                                     Light_Guard_Bypass=>"Light_Guard_Bypass(1)",
                                     System_Busy:="System_1_Busy");
                100401:
                    "Feed_BCNV_Cnv1(1)"( System_No := 1,
                                     Level := 4,
                                     Light_Guard_IO:="LIGHT GUARDS C1101 - CH1",
                                     Light_Guard_Bypass=>"Light_Guard_Bypass(1)",
                                     System_Busy:="System_1_Busy");
                100501:
                    "Feed_BCNV_Cnv1(1)"( System_No := 1,
                                     Level := 5,
                                     Light_Guard_IO:="LIGHT GUARDS C1101 - CH1",
                                     Light_Guard_Bypass=>"Light_Guard_Bypass(1)",
                                     System_Busy:="System_1_Busy");
                100601:
                    "Feed_BCNV_Cnv1(1)"( System_No := 1,
                                     Level := 6,
                                     Light_Guard_IO:="LIGHT GUARDS C1101 - CH1",
                                     Light_Guard_Bypass=>"Light_Guard_Bypass(1)",
                                     System_Busy:="System_1_Busy");
                100701:
                    "Feed_BCNV_Cnv1(1)"( System_No := 1,
                                     Level := 7,
                                     Light_Guard_IO:="LIGHT GUARDS C1101 - CH1",
                                     Light_Guard_Bypass=>"Light_Guard_Bypass(1)",
                                     System_Busy:="System_1_Busy");
                100801:
                    "Feed_BCNV_Cnv1(1)"( System_No := 1,
                                     Level := 8,
                                     Light_Guard_IO:="LIGHT GUARDS C1101 - CH1",
                                     Light_Guard_Bypass=>"Light_Guard_Bypass(1)",
                                     System_Busy:="System_1_Busy");
                    //CNV 2
                110101:
                    "Feed_BCNV_Cnv2(1)"( System_No := 1,
                                     Level := 1,
                                     Light_Guard_IO:="LIGHT GUARDS C1201 - CH1",
                                     Light_Guard_Bypass=>"Light_Guard_Bypass(1)",
                                     System_Busy:="System_1_Busy");
                110201:
                    "Feed_BCNV_Cnv2(1)"( System_No := 1,
                                     Level := 2,
                                     Light_Guard_IO:="LIGHT GUARDS C1201 - CH1",
                                     Light_Guard_Bypass=>"Light_Guard_Bypass(1)",
                                     System_Busy:="System_1_Busy");
                110301:
                    "Feed_BCNV_Cnv2(1)"( System_No := 1,
                                     Level := 3,
                                     Light_Guard_IO:="LIGHT GUARDS C1201 - CH1",
                                     Light_Guard_Bypass=>"Light_Guard_Bypass(1)",
                                     System_Busy:="System_1_Busy");
                110401:
                    "Feed_BCNV_Cnv2(1)"( System_No := 1,
                                     Level := 4,
                                     Light_Guard_IO:="LIGHT GUARDS C1201 - CH1",
                                     Light_Guard_Bypass=>"Light_Guard_Bypass(1)",
                                     System_Busy:="System_1_Busy");
                110501:
                    "Feed_BCNV_Cnv2(1)"( System_No := 1,
                                     Level := 5,
                                     Light_Guard_IO:="LIGHT GUARDS C1201 - CH1",
                                     Light_Guard_Bypass=>"Light_Guard_Bypass(1)",
                                     System_Busy:="System_1_Busy");
                110601:
                    "Feed_BCNV_Cnv2(1)"( System_No := 1,
                                     Level := 6,
                                     Light_Guard_IO:="LIGHT GUARDS C1201 - CH1",
                                     Light_Guard_Bypass=>"Light_Guard_Bypass(1)",
                                     System_Busy:="System_1_Busy");
                110701:
                    "Feed_BCNV_Cnv2(1)"( System_No := 1,
                                     Level := 7,
                                     Light_Guard_IO:="LIGHT GUARDS C1201 - CH1",
                                     Light_Guard_Bypass=>"Light_Guard_Bypass(1)",
                                     System_Busy:="System_1_Busy");
                110801:
                    "Feed_BCNV_Cnv2(1)"( System_No := 1,
                                     Level := 8,
                                     Light_Guard_IO:="LIGHT GUARDS C1201 - CH1",
                                     Light_Guard_Bypass=>"Light_Guard_Bypass(1)",
                                     System_Busy:="System_1_Busy");
                    //SYSTEM 2
                    //CNV 1
                100102:
                    "Feed_BCNV_Cnv1(1)"(System_No := 2,
                                        Level := 1,
                                        Light_Guard_IO := "LIGHT GUARDS C2101 - CH1",
                                        Light_Guard_Bypass=>"Light_Guard_Bypass(2)",
                                        System_Busy := "System_2_Busy");
                100202:
                    "Feed_BCNV_Cnv1(1)"( System_No := 2,
                                     Level := 2,
                                     Light_Guard_IO:="LIGHT GUARDS C2101 - CH1",
                                     Light_Guard_Bypass=>"Light_Guard_Bypass(2)",
                                     System_Busy:="System_2_Busy");
                100302:
                    "Feed_BCNV_Cnv1(1)"( System_No := 2,
                                     Level := 3,
                                     Light_Guard_IO:="LIGHT GUARDS C2101 - CH1",
                                     Light_Guard_Bypass=>"Light_Guard_Bypass(2)",
                                     System_Busy:="System_2_Busy");
                100402:
                    "Feed_BCNV_Cnv1(1)"( System_No := 2,
                                     Level := 4,
                                     Light_Guard_IO:="LIGHT GUARDS C2101 - CH1",
                                     Light_Guard_Bypass=>"Light_Guard_Bypass(2)",
                                     System_Busy:="System_2_Busy");
                100502:
                    "Feed_BCNV_Cnv1(1)"( System_No := 2,
                                     Level := 5,
                                     Light_Guard_IO:="LIGHT GUARDS C2101 - CH1",
                                     Light_Guard_Bypass=>"Light_Guard_Bypass(2)",
                                     System_Busy:="System_2_Busy");
                100602:
                    "Feed_BCNV_Cnv1(1)"( System_No := 2,
                                     Level := 6,
                                     Light_Guard_IO:="LIGHT GUARDS C2101 - CH1",
                                     Light_Guard_Bypass=>"Light_Guard_Bypass(2)",
                                     System_Busy:="System_2_Busy");
                100702:
                    "Feed_BCNV_Cnv1(1)"( System_No := 2,
                                     Level := 7,
                                     Light_Guard_IO:="LIGHT GUARDS C2101 - CH1",
                                     Light_Guard_Bypass=>"Light_Guard_Bypass(2)",
                                     System_Busy:="System_2_Busy");
                100802:
                    "Feed_BCNV_Cnv1(1)"( System_No := 2,
                                     Level := 8,
                                     Light_Guard_IO:="LIGHT GUARDS C2101 - CH1",
                                     Light_Guard_Bypass=>"Light_Guard_Bypass(2)",
                                     System_Busy:="System_2_Busy");
                    //CNV 2
                110102:
                    "Feed_BCNV_Cnv2(1)"( System_No := 2,
                                     Level := 1,
                                     Light_Guard_IO:="LIGHT GUARDS C2201 - CH1",
                                     Light_Guard_Bypass=>"Light_Guard_Bypass(2)",
                                     System_Busy:="System_2_Busy");
                110202:
                    "Feed_BCNV_Cnv2(1)"( System_No := 2,
                                     Level := 2,
                                     Light_Guard_IO:="LIGHT GUARDS C2201 - CH1",
                                     Light_Guard_Bypass=>"Light_Guard_Bypass(2)",
                                     System_Busy:="System_2_Busy");
                110302:
                    "Feed_BCNV_Cnv2(1)"( System_No := 2,
                                     Level := 3,
                                     Light_Guard_IO:="LIGHT GUARDS C2201 - CH1",
                                     Light_Guard_Bypass=>"Light_Guard_Bypass(2)",
                                     System_Busy:="System_2_Busy");
                110402:
                    "Feed_BCNV_Cnv2(1)"( System_No := 2,
                                     Level := 4,
                                     Light_Guard_IO:="LIGHT GUARDS C2201 - CH1",
                                     Light_Guard_Bypass=>"Light_Guard_Bypass(2)",
                                     System_Busy:="System_2_Busy");
                110502:
                    "Feed_BCNV_Cnv2(1)"( System_No := 2,
                                     Level := 5,
                                     Light_Guard_IO:="LIGHT GUARDS C2201 - CH1",
                                     Light_Guard_Bypass=>"Light_Guard_Bypass(2)",
                                     System_Busy:="System_2_Busy");
                110602:
                    "Feed_BCNV_Cnv2(1)"( System_No := 2,
                                     Level := 6,
                                     Light_Guard_IO:="LIGHT GUARDS C2201 - CH1",
                                     Light_Guard_Bypass=>"Light_Guard_Bypass(2)",
                                     System_Busy:="System_2_Busy");
                110702:
                    "Feed_BCNV_Cnv2(1)"( System_No := 2,
                                     Level := 7,
                                     Light_Guard_IO:="LIGHT GUARDS C2201 - CH1",
                                     Light_Guard_Bypass=>"Light_Guard_Bypass(2)",
                                     System_Busy:="System_2_Busy");
                110802:
                    "Feed_BCNV_Cnv2(1)"( System_No := 2,
                                     Level := 8,
                                     Light_Guard_IO:="LIGHT GUARDS C2201 - CH1",
                                     Light_Guard_Bypass=>"Light_Guard_Bypass(2)",
                                     System_Busy:="System_2_Busy");
                    //SYSTEM 3
                    //CNV 1
                100103:
                    "Feed_BCNV_Cnv1(1)"( System_No := 3,
                                     Level := 1,
                                     Light_Guard_IO:="LIGHT GUARDS C3101 - CH1",
                                     Light_Guard_Bypass=>"Light_Guard_Bypass(3)",
                                     System_Busy:="System_3_Busy");
                100203:
                    "Feed_BCNV_Cnv1(1)"( System_No := 3,
                                     Level := 2,
                                     Light_Guard_IO:="LIGHT GUARDS C3101 - CH1",
                                     Light_Guard_Bypass=>"Light_Guard_Bypass(3)",
                                     System_Busy:="System_3_Busy");
                100303:
                    "Feed_BCNV_Cnv1(1)"( System_No := 3,
                                     Level := 3,
                                     Light_Guard_IO:="LIGHT GUARDS C3101 - CH1",
                                     Light_Guard_Bypass=>"Light_Guard_Bypass(3)",
                                     System_Busy:="System_3_Busy");
                100403:
                    "Feed_BCNV_Cnv1(1)"( System_No := 3,
                                     Level := 4,
                                     Light_Guard_IO:="LIGHT GUARDS C3101 - CH1",
                                     Light_Guard_Bypass=>"Light_Guard_Bypass(3)",
                                     System_Busy:="System_3_Busy");
                100503:
                    "Feed_BCNV_Cnv1(1)"( System_No := 3,
                                     Level := 5,
                                     Light_Guard_IO:="LIGHT GUARDS C3101 - CH1",
                                     Light_Guard_Bypass=>"Light_Guard_Bypass(3)",
                                     System_Busy:="System_3_Busy");
                100603:
                    "Feed_BCNV_Cnv1(1)"( System_No := 3,
                                     Level := 6,
                                     Light_Guard_IO:="LIGHT GUARDS C3101 - CH1",
                                     Light_Guard_Bypass=>"Light_Guard_Bypass(3)",
                                     System_Busy:="System_3_Busy");
                100703:
                    "Feed_BCNV_Cnv1(1)"( System_No := 3,
                                     Level := 7,
                                     Light_Guard_IO:="LIGHT GUARDS C3101 - CH1",
                                     Light_Guard_Bypass=>"Light_Guard_Bypass(3)",
                                     System_Busy:="System_3_Busy");
                100803:
                    "Feed_BCNV_Cnv1(1)"( System_No := 3,
                                     Level := 8,
                                     Light_Guard_IO:="LIGHT GUARDS C3101 - CH1",
                                     Light_Guard_Bypass=>"Light_Guard_Bypass(3)",
                                     System_Busy:="System_3_Busy");
                    //CNV 2
                110103:
                    "Feed_BCNV_Cnv2(1)"( System_No := 3,
                                     Level := 1,
                                     Light_Guard_IO:="LIGHT GUARDS C3201 - CH1",
                                     Light_Guard_Bypass=>"Light_Guard_Bypass(3)",
                                     System_Busy:="System_3_Busy");
                110203:
                    "Feed_BCNV_Cnv2(1)"( System_No := 3,
                                     Level := 2,
                                     Light_Guard_IO:="LIGHT GUARDS C3201 - CH1",
                                     Light_Guard_Bypass=>"Light_Guard_Bypass(3)",
                                     System_Busy:="System_3_Busy");
                110303:
                    "Feed_BCNV_Cnv2(1)"( System_No := 3,
                                     Level := 3,
                                     Light_Guard_IO:="LIGHT GUARDS C3201 - CH1",
                                     Light_Guard_Bypass=>"Light_Guard_Bypass(3)",
                                     System_Busy:="System_3_Busy");
                110403:
                    "Feed_BCNV_Cnv2(1)"( System_No := 3,
                                     Level := 4,
                                     Light_Guard_IO:="LIGHT GUARDS C3201 - CH1",
                                     Light_Guard_Bypass=>"Light_Guard_Bypass(3)",
                                     System_Busy:="System_3_Busy");
                110503:
                    "Feed_BCNV_Cnv2(1)"( System_No := 3,
                                     Level := 5,
                                     Light_Guard_IO:="LIGHT GUARDS C3201 - CH1",
                                     Light_Guard_Bypass=>"Light_Guard_Bypass(3)",
                                     System_Busy:="System_3_Busy");
                110603:
                    "Feed_BCNV_Cnv2(1)"( System_No := 3,
                                     Level := 6,
                                     Light_Guard_IO:="LIGHT GUARDS C3201 - CH1",
                                     Light_Guard_Bypass=>"Light_Guard_Bypass(3)",
                                     System_Busy:="System_3_Busy");
                110703:
                    "Feed_BCNV_Cnv2(1)"( System_No := 3,
                                     Level := 7,
                                     Light_Guard_IO:="LIGHT GUARDS C3201 - CH1",
                                     Light_Guard_Bypass=>"Light_Guard_Bypass(3)",
                                     System_Busy:="System_3_Busy");
                110803:
                    "Feed_BCNV_Cnv2(1)"( System_No := 3,
                                     Level := 8,
                                     Light_Guard_IO:="LIGHT GUARDS C3201 - CH1",
                                     Light_Guard_Bypass=>"Light_Guard_Bypass(3)",
                                     System_Busy:="System_3_Busy");
                    //SYSTEM 4
                    //CNV 2
                100104:
                    "Feed_BCNV_Cnv1(1)"( System_No := 4,
                                     Level := 1,
                                     Light_Guard_IO:=TRUE,
                                     Light_Guard_Bypass=>#No_Light_Guard,
                                     System_Busy:="System_4_Busy");
                100204:
                    "Feed_BCNV_Cnv1(1)"( System_No := 4,
                                     Level := 2,
                                     Light_Guard_IO:=TRUE,
                                     Light_Guard_Bypass=>#No_Light_Guard,
                                     System_Busy:="System_4_Busy");
                100304:
                    "Feed_BCNV_Cnv1(1)"( System_No := 4,
                                     Level := 3,
                                     Light_Guard_IO:=TRUE,
                                     Light_Guard_Bypass=>#No_Light_Guard,
                                     System_Busy:="System_4_Busy");
                100404:
                    "Feed_BCNV_Cnv1(1)"( System_No := 4,
                                     Level := 4,
                                     Light_Guard_IO:=TRUE,
                                     Light_Guard_Bypass=>#No_Light_Guard,
                                     System_Busy:="System_4_Busy");
                100504:
                    "Feed_BCNV_Cnv1(1)"( System_No := 4,
                                     Level := 5,
                                     Light_Guard_IO:=TRUE,
                                     Light_Guard_Bypass=>#No_Light_Guard,
                                     System_Busy:="System_4_Busy");
                100604:
                    "Feed_BCNV_Cnv1(1)"( System_No := 4,
                                     Level := 6,
                                     Light_Guard_IO:=TRUE,
                                     Light_Guard_Bypass=>#No_Light_Guard,
                                     System_Busy:="System_4_Busy");
                100704:
                    "Feed_BCNV_Cnv1(1)"( System_No := 4,
                                     Level := 7,
                                     Light_Guard_IO:=TRUE,
                                     Light_Guard_Bypass=>#No_Light_Guard,
                                     System_Busy:="System_4_Busy");
                100804:
                    "Feed_BCNV_Cnv1(1)"( System_No := 4,
                                     Level := 8,
                                     Light_Guard_IO:=TRUE,
                                     Light_Guard_Bypass=>#No_Light_Guard,
                                     System_Busy:="System_4_Busy");
                    //SYSTEM 5
                120005:
                    "Feed_ECNV(1)"( System_No := 5);
                    //CNV 2
                100105:
                    "Feed_BCNV_Cnv1(1)"( System_No := 5,
                                     Level := 1,
                                     Light_Guard_IO:=TRUE,
                                     Light_Guard_Bypass=>#No_Light_Guard,
                                     System_Busy:="System_5_Busy");
                100205:
                    "Feed_BCNV_Cnv1(1)"( System_No := 5,
                                     Level := 2,
                                     Light_Guard_IO:=TRUE,
                                     Light_Guard_Bypass=>#No_Light_Guard,
                                     System_Busy:="System_5_Busy");
                100305:
                    "Feed_BCNV_Cnv1(1)"( System_No := 5,
                                     Level := 3,
                                     Light_Guard_IO:=TRUE,
                                     Light_Guard_Bypass=>#No_Light_Guard,
                                     System_Busy:="System_5_Busy");
                100405:
                    "Feed_BCNV_Cnv1(1)"( System_No := 5,
                                     Level := 4,
                                     Light_Guard_IO:=TRUE,
                                     Light_Guard_Bypass=>#No_Light_Guard,
                                     System_Busy:="System_5_Busy");
                100505:
                    "Feed_BCNV_Cnv1(1)"( System_No := 5,
                                     Level := 5,
                                     Light_Guard_IO:=TRUE,
                                     Light_Guard_Bypass=>#No_Light_Guard,
                                     System_Busy:="System_5_Busy");
                100605:
                    "Feed_BCNV_Cnv1(1)"( System_No := 5,
                                     Level := 6,
                                     Light_Guard_IO:=TRUE,
                                     Light_Guard_Bypass=>#No_Light_Guard,
                                     System_Busy:="System_5_Busy");
                100705:
                    "Feed_BCNV_Cnv1(1)"( System_No := 5,
                                     Level := 7,
                                     Light_Guard_IO:=TRUE,
                                     Light_Guard_Bypass=>#No_Light_Guard,
                                     System_Busy:="System_5_Busy");
                100805:
                    "Feed_BCNV_Cnv1(1)"( System_No := 5,
                                     Level := 8,
                                     Light_Guard_IO:=TRUE,
                                     Light_Guard_Bypass=>#No_Light_Guard,
                                     System_Busy:="System_5_Busy");
            END_CASE;
        END_IF;
    END_REGION
END_REGION


//RESET CHARGE BITS
#T_Reset_Charge.TON(IN := "Screen_DB".Charge_VTD OR "Screen_DB".Charge_Cnv OR "Screen_DB".Charge_VTD_Commands OR "Screen_DB".Charge_Cnv_Commands,
                       PT := T#2S);

   IF #T_Reset_Charge.Q THEN
    "Screen_DB".Charge_VTD := FALSE;
    "Screen_DB".Charge_Cnv := FALSE;
    "Screen_DB".Charge_VTD_Commands := FALSE;
    "Screen_DB".Charge_Cnv_Commands := FALSE;
END_IF;

END_FUNCTION_BLOCK